// TIA Portal V21 export
// export: Created 2026-11-10T07:35:23.821205Z, ExportSetting WithDefaults, DisplayName Totally Integrated Automation Portal, DisplayVersion V21 Update 3, DisplayName STEP 7 Professional, DisplayVersion V21 Update 3, DisplayName STEP 7 Safety, DisplayVersion V21, DisplayName Tech WebApplication, DisplayVersion V21, DisplayName WinCC Basic/Comfort/Advanced, DisplayVersion V21 Update 3, DisplayName WinCC Unified, DisplayVersion V21 Update 3
FUNCTION_BLOCK "FB_Lad_ex157"   // FB59, LAD
{ S7_Optimized_Access := 'TRUE' }
VERSION : 0.1
// stored: AutoNumber true, IsIECCheckEnabled false, IsRetainMemResEnabled false, MemoryReserve 100, SetENOAutomatically false, UDAEnableTagReadback false
   VAR_INPUT
      v_master : Int;
      v_station : Int;
      v_slot : Int;
      v_subslot : Int;
      v_ret_val : Int;
   END_VAR
   VAR_OUTPUT
      v_laddr : HW_IO;
   END_VAR
BEGIN

REGION Network 1: GEO_LOG - Determine hardware identifier from slot
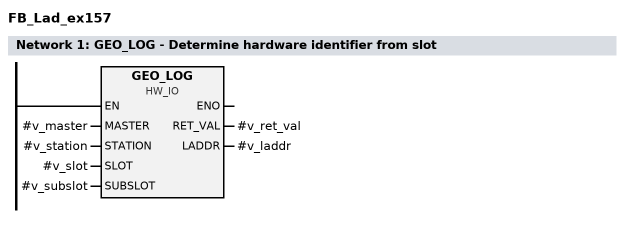
   RUNG wire#powerrail
      { S7_Templates := "laddr_type := HW_IO" } GEO_LOG(MASTER := #v_master, STATION := #v_station, SLOT := #v_slot, SUBSLOT := #v_subslot, RET_VAL => #v_ret_val, LADDR => #v_laddr)
   END_RUNG
   // the same network as SCL:
   #v_ret_val := GEO_LOG(MASTER := #v_master,
                         STATION := #v_station,
                         SLOT := #v_slot,
                         SUBSLOT := #v_subslot,
                         LADDR => #v_laddr);
END_REGION
END_FUNCTION_BLOCK
